Fanuc KAREL source: kt00646.KL

-- PROVISIONAL review KL for V1013-1; original PC SHA256 48af6d36c95c8cf6c8008cf071107fd9f670ad70d786b0beb8665354ed987a1f
-- Incomplete behavior may be omitted. Consult companion uncertainty JSON. Do not deploy.
PROGRAM KT00646
%NOLOCKGROUP
VAR
  OUT : INTEGER
-- UNRESOLVED_DECL H1 type=002017
-- UNRESOLVED_DECL H2 type=002017
BEGIN
  -- UNRESOLVED_PC offsets 5-19; opcodes 2E,22,9D,33,B4
  -- UNRESOLVED_PC offsets 24-38; opcodes 2E,22,9D,33,B4
  -- UNRESOLVED_PC offsets 43-57; opcodes 2E,22,9D,33,B4
  -- UNRESOLVED_PC offsets 62-76; opcodes 2E,22,9D,33,B4
  -- UNRESOLVED_PC offsets 81-96; opcodes 22,9D,33,B3,23
  -- UNRESOLVED_PC offsets 101-105; opcodes 7F
END KT00646
